Staubli VAL3: _systemStates.pgx

public program _systemStates()
begin
  // while true
  //程序运行中
  rs:bIsCycle=(taskStatus("cycle")>-1)
  //home
  rs:bIsHome=(abs(herej()-saveData:jHome)<{2,2,2,2,2,2})
  //使能上电
  rs:bPowerON=(isPowered()==true)
  //远程模式
  rs:bIsRemoteAuto=(workingMode()==4)
  //机器人正在移动
  rs:bIsMoving=(isSettled()==false)
  //机器人急停
  rs:bIsEstop=(esStatus()!=0)
  //
  rs:bIsReady=!rs:bIsCycle and rs:bIsHome and rs:bPowerON and !rs:bIsEstop and  rs:bIsRemoteAuto
  //程序报错
  rs:bIsError=(taskStatus("cycle")>1)

  // delay(0)
  // endWhile

end
